(* IEC 61131-3 sources: garage-sweeper/PLC/src/Adapters/Simulation, 5 files *)

(* ---- Accelerometer_Simulated.st ---- *)
{attribute 'linkalways'}
{attribute 'no_explicit_call' := 'Use the methods of this class'}
{attribute 'enable_dynamic_creation'}
FUNCTION_BLOCK Accelerometer_Simulated IMPLEMENTS I_Accelerometer
VAR
	link : REFERENCE TO SimulatorLink;
END_VAR
METHOD FB_init : BOOL
VAR_INPUT
	bInitRetains : BOOL;
	bInCopyCode : BOOL;
	simulator : REFERENCE TO SimulatorLink;
END_VAR
// @impl
link REF= simulator;
END_METHOD
PROPERTY AccelerationInMPerS2 : Vector3
GET
AccelerationInMPerS2 := SimulatorIo.feedback.accelerationInMPerS2;
END_GET
END_PROPERTY
PROPERTY TimestampInNs : ULINT
GET
TimestampInNs := SimulatorIo.feedback.timeInNs;
END_GET
END_PROPERTY
PROPERTY IsValid : BOOL
GET
IsValid := __ISVALIDREF(link) AND_THEN link.IsConnected;
END_GET
END_PROPERTY

(* ---- DigitalOut_SimulatedLidarPower.st ---- *)
{attribute 'linkalways'}
{attribute 'no_explicit_call' := 'Use the methods of this class'}
{attribute 'enable_dynamic_creation'}
FUNCTION_BLOCK DigitalOut_SimulatedLidarPower IMPLEMENTS I_DigitalOut
METHOD SwitchOn
// @impl
SimulatorIo.command.isLidarPowered := TRUE;
END_METHOD
METHOD SwitchOff
// @impl
SimulatorIo.command.isLidarPowered := FALSE;
END_METHOD
PROPERTY IsOn : BOOL
GET
IsOn := SimulatorIo.command.isLidarPowered;
END_GET
END_PROPERTY

(* ---- Gyro_Simulated.st ---- *)
{attribute 'linkalways'}
{attribute 'no_explicit_call' := 'Use the methods of this class'}
{attribute 'enable_dynamic_creation'}
FUNCTION_BLOCK Gyro_Simulated IMPLEMENTS I_Gyro
VAR
	link : REFERENCE TO SimulatorLink;
END_VAR
METHOD FB_init : BOOL
VAR_INPUT
	bInitRetains : BOOL;
	bInCopyCode : BOOL;
	simulator : REFERENCE TO SimulatorLink;
END_VAR
// @impl
link REF= simulator;
END_METHOD
METHOD StartBiasCalibration
// @impl
// The simulated gyro has no calibration of its own. Bias is estimated in HeadingFusion.
END_METHOD
PROPERTY YawRateInRadPerS : LREAL
GET
YawRateInRadPerS := SimulatorIo.feedback.angularRateInRadPerS.z;
END_GET
END_PROPERTY
PROPERTY AngularRateInRadPerS : Vector3
GET
AngularRateInRadPerS := SimulatorIo.feedback.angularRateInRadPerS;
END_GET
END_PROPERTY
PROPERTY TimestampInNs : ULINT
GET
TimestampInNs := SimulatorIo.feedback.timeInNs;
END_GET
END_PROPERTY
PROPERTY IsValid : BOOL
GET
IsValid := __ISVALIDREF(link) AND_THEN link.IsConnected;
END_GET
END_PROPERTY

(* ---- Lidar_Simulated.st ---- *)
{attribute 'linkalways'}
{attribute 'no_explicit_call' := 'Use the methods of this class'}
{attribute 'enable_dynamic_creation'}
FUNCTION_BLOCK Lidar_Simulated IMPLEMENTS I_Lidar
VAR
	notConnectedError : HardwareError := (isActive := TRUE, id := Constants.SIMULATOR_NOT_CONNECTED_ERROR_ID, text := 'Simulatoren er ikke tilkoblet');
	link : REFERENCE TO SimulatorLink;
	_isRunning : BOOL;
	lastSequence : UDINT;
END_VAR
METHOD FB_init : BOOL
VAR_INPUT
	bInitRetains : BOOL;
	bInCopyCode : BOOL;
	simulator : REFERENCE TO SimulatorLink;
END_VAR
// @impl
link REF= simulator;
END_METHOD
METHOD Start
// @impl
_isRunning := TRUE;
lastSequence := SimulatorIo.scan.sequence;
END_METHOD
METHOD Stop
// @impl
_isRunning := FALSE;
END_METHOD
METHOD TryGetScan : BOOL
VAR_INPUT
	scan : REFERENCE TO LaserScan;
END_VAR
// @impl
IF NOT _isRunning OR_ELSE SimulatorIo.scan.sequence = lastSequence THEN
	RETURN;
END_IF
lastSequence := SimulatorIo.scan.sequence;
scan := SimulatorIo.scan;
TryGetScan := TRUE;
END_METHOD
PROPERTY IsRunning : BOOL
GET
IsRunning := _isRunning;
END_GET
END_PROPERTY
PROPERTY Error : HardwareError
GET
IF NOT __ISVALIDREF(link) OR_ELSE NOT link.IsConnected THEN
	Error := notConnectedError;
END_IF
END_GET
END_PROPERTY

(* ---- SimulatorLink.st ---- *)
{attribute 'linkalways'}
{attribute 'no_explicit_call' := 'Use the methods of this class'}
{attribute 'enable_dynamic_creation'}
FUNCTION_BLOCK SimulatorLink
VAR
	cycle : UDINT;
	lastSequence : UDINT;
	silentCycles : UDINT;
	_isConnected : BOOL;
END_VAR
METHOD Execute
// @impl
cycle := cycle + 1;
SimulatorIo.command.version := Constants.SIMULATOR_PROTOCOL_VERSION;
SimulatorIo.command.cycle := cycle;
SimulatorIo.command.plcTimeInNs := F_GetSystemTime() * 100;

IF SimulatorIo.feedback.sequence <> lastSequence THEN
	lastSequence := SimulatorIo.feedback.sequence;
	silentCycles := 0;
ELSIF silentCycles < Constants.SIMULATOR_TIMEOUT_IN_CYCLES THEN
	silentCycles := silentCycles + 1;
END_IF

_isConnected := SimulatorIo.feedback.version = Constants.SIMULATOR_PROTOCOL_VERSION
	AND silentCycles < Constants.SIMULATOR_TIMEOUT_IN_CYCLES;
END_METHOD
PROPERTY IsConnected : BOOL
GET
IsConnected := _isConnected;
END_GET
END_PROPERTY
